(* PLC project v0.6.03_RunVisu.project, CODESYS CODESYS V3.5 SP19 Patch 1 *)
(* stored: creationDateTime 2026-08-15T01:10:37.9768184, modificationDateTime 2026-08-14T23:30:12.3399581 *)

(* ═══════════════════════════════════════════════════════════════ 📤 PRG_06_Outputs_LD — Écriture des SORTIES physiques (PROGRAMME LADDER) ─────────────────────────────────────────────────────────────── 📄 Doc : DOC/AF/AF_Partie-06_Acquisition_Qualification_IO_v2.3.md §5 ⚙️ Exécuté par la tâche PLC en position 6 (après PRG_05_Translation). 📄 Converti automatiquement en Ladder Diagram (<LD>) dans CODESYS. 🛡️ LOT_STRUCTURE_INTERLOCKS_LD (2026-08) : barrières finales M1/M2/M3 rendues visibles — FB_WinchOutputInterlock_LD (×2) et FB_TranslationOutputInterlock_LD (×1) câblés en amont des coils, contacts nommés sur variables qualifiées (visibilité maintenance : interlocks/safety qui coupent chaque actionneur lisibles directement dans le réseau Ladder, sans ouvrir un autre POU). 🔒 SafetyStructureNotValidated reste TRUE : AUCUNE sortie physique moteur/frein n'est autorisée tant que ce garde-fou n'est pas retiré dans un lot safety validé séparément (voir alerte ci-dessous). ⚠️ Écart connu, HORS PÉRIMÈTRE de ce lot (signalé, pas corrigé ici) : FB_Safety_Winch / FB_Safety_Translation (7 mécanismes Méca A→E, PowerCutOff métier) ne sont appelés nulle part dans CODE/ à ce jour. ST_WinchFinalInterlockRequest / ST_TranslationFinalInterlockRequest ne portent donc que SafeStop (partiel) — voir PLAN_TASK lot "5 Reliquats safety" (T72-T74). Ce lot ne câble que ce qui existe déjà en amont ; ne pas déduire que la safety métier complète est active. 🗑️ FB_Output retiré (2026-08) : inverseur pur (State := Command XOR InvertLogic) jamais utilisé avec InvertLogic <> FALSE (REX 2026-08-04, feedback déjà retiré). Coils câblées directement sur les sorties des interlocks finaux — élimine 15 blocs sans valeur ajoutée et simplifie la lecture maintenance. 🆕 LOT2 (2026-08-05) : sortie moteur AC600 M3 raccordée. DriveControlWord (mot commande 0x3101) et DriveFreqRefWord (consigne fréquence WORD, registre 0x3100, échelle ×100 confirmée terrain — WORD 5000 = 50,00 Hz) capturés en variables locales M3_DriveControlWord / M3_DriveFreqRefWord. Mapping E/S CODESYS (Device.export) manuel restant — voir §2 ci-dessous. ═══════════════════════════════════════════════════════════════ *)
PROGRAM PRG_06_Outputs_LD_1
  VAR_OUTPUT
    EmergencyArmingPulseActive : BOOL;  (* 🐛 FIX 2026-08-05 (confirmé câblé réel par l'utilisateur) : PowerKeepAlive_A_RQ/ PowerKeepAlive_B_RQ/EmergencyArming_RQ retirés d'ici — même collision de portée que M1/M2/M3 (voir §2). Cibles renommées : PowerKeepAliveACmd/BCmd/ EmergencyArmingCmd, déclarées en VAR locale ci-dessous. *)
    EmergencyArmingLockoutActive : BOOL;
    ArmingSeqStep : INT;
    RedundancyTestFailed : BOOL;
    EmergencyArmingFailed : BOOL;
    EmergencyState : ST_Safety_Emergency_State;
    EmergencyDiag : ST_Safety_Emergency_Diag;
    PowerCutOffActive : BOOL;  (* TRUE = demande de coupure finale active *)
    SafetyStructureNotValidated : BOOL := FALSE;  (* 🔓 Garde-fou désactivé : les autorisations M1/M2/M3 sont liées dynamiquement à leurs sécurités *)
    M1InterlockEnable : BOOL;  (* 🔧 FIX 2026-08-14 (audit sécurité) : Enable ne coupe plus que sur PowerCutOff (barrière finale, AF02 §2, AF06 §5 "SafeStop laisse la décélération métier se terminer"). SafeStop/ Error retirés du calcul — SafeStop est une rampe rapide gérée en amont par FB_Winch/ FB_Translation (Enable maintenu, AGENTS.md, TC-P03-001) ; Error mirait tout ErrorId y compris les mécanismes SafeStop-only, donc coupait Enable pour la même mauvaise raison. Couper ici sur SafeStop/Error écrasait la rampe déjà calculée en amont en un arrêt brutal — contraire à la doctrine Enable>SafeStop>StartStop. Gate finale M1 : WinchM1FinalInterlockRequest.Enable AND NOT WinchM1FinalInterlockRequest.PowerCutOff *)
    M2InterlockEnable : BOOL;  (* Gate finale M2 : WinchM2FinalInterlockRequest.Enable AND NOT WinchM2FinalInterlockRequest.PowerCutOff *)
    M3InterlockEnable : BOOL;  (* Gate finale M3 : TranslationFinalInterlockRequest.Enable AND NOT TranslationFinalInterlockRequest.PowerCutOff *)
    M1BlockedBySafetyInfo : BOOL;  (* 🆕 Réseau informatif séparé (demande utilisateur) : visibilité maintenance de ce qui bloque (SafeStop/Error), SANS influencer Enable — juste de l'information en Watch/Ladder. *)
    M2BlockedBySafetyInfo : BOOL;
    M3BlockedBySafetyInfo : BOOL;
    TranslationBrakeCmd : BOOL;  (* 🐛 FIX 2026-08-05 : les noms Device bruts ( *_DQ / *_RQ ), ex. M1_RelayFwd_Up_DQ, M3_BrakeRelease_RQ) NE SONT PLUS déclarés ici — les déclarer créait une collision de portée avec la variable GLOBALE homonyme créée par le mapping E/S CODESYS (Device.export), qui masquait silencieusement le pilotage matériel réel (voir §2 plus bas pour le détail et la liste des chemins qualifiés à mapper). Demande frein M3 arbitrée — cible du mapping E/S *)
    M3_DriveControlWord : WORD;  (* Mot de commande variateur M3 (0x3101) — cible du mapping E/S *)
    M3_DriveFreqRefWord : WORD;  (* Consigne fréquence variateur M3 (0x3100, x100) — cible du mapping E/S *)
  END_VAR
  VAR
    instWinchOutputInterlockM1 : FB_WinchOutputInterlock_LD;
    instWinchOutputInterlockM2 : FB_WinchOutputInterlock_LD;
    instTranslationOutputInterlockM3 : FB_TranslationOutputInterlock_LD;
    M1RelayFwd : BOOL;
    M1RelayRev : BOOL;
    M1SpeedContactor1 : BOOL;
    M1SpeedContactor2 : BOOL;
    M1SpeedContactor3 : BOOL;
    M1SpeedContactor4 : BOOL;
    M1BrakeCmd : BOOL;
    M2RelayFwd : BOOL;
    M2RelayRev : BOOL;
    M2SpeedContactor1 : BOOL;
    M2SpeedContactor2 : BOOL;
    M2SpeedContactor3 : BOOL;
    M2SpeedContactor4 : BOOL;
    M2BrakeCmd : BOOL;
    KoboldContactorCmd : BOOL;
    PowerCutOffReq : BOOL;
    PowerKeepAliveACmd : BOOL;  (* Maintien puissance voie A — cible du mapping E/S *)
    PowerKeepAliveBCmd : BOOL;  (* Maintien puissance voie B — cible du mapping E/S *)
    EmergencyArmingCmd : BOOL;  (* Impulsion réarmement — cible du mapping E/S *)
    instSafetyEmergencyManagement : FB_Safety_EmergencyManagement;
  END_VAR

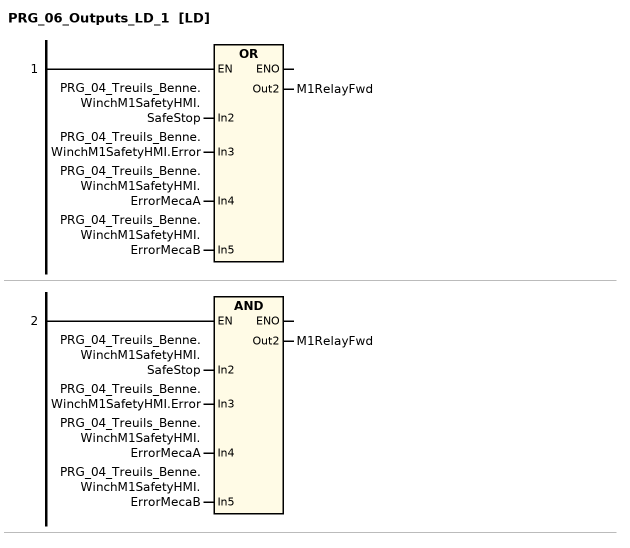
(* LD diagram, written out as Structured Text *)

M1RelayFwd := PRG_04_Treuils_Benne.WinchM1SafetyHMI.SafeStop OR PRG_04_Treuils_Benne.WinchM1SafetyHMI.Error OR PRG_04_Treuils_Benne.WinchM1SafetyHMI.ErrorMecaA OR PRG_04_Treuils_Benne.WinchM1SafetyHMI.ErrorMecaB;

M1RelayFwd := PRG_04_Treuils_Benne.WinchM1SafetyHMI.SafeStop AND PRG_04_Treuils_Benne.WinchM1SafetyHMI.Error AND PRG_04_Treuils_Benne.WinchM1SafetyHMI.ErrorMecaA AND PRG_04_Treuils_Benne.WinchM1SafetyHMI.ErrorMecaB;
END_PROGRAM
